// Pools d'objets (docs/04 § 9) : instances déclarées une fois pour toutes, attribuées au déploiement par
// FB_ObjectFactory. La bibliothèque fournit FB_DefaultPools ; un projet peut donner les siens.
INTERFACE I_ObjectPools

// Nombre d'éléments du pool d'un type, 0 = type absent
METHOD PoolSize : UINT
VAR_INPUT
    nType : UINT;
END_VAR
END_METHOD

// N° du pool d'un type : deux types qui partagent un pool (axe linéaire et rotatif, modules) ont le même n°
METHOD PoolId : UINT
VAR_INPUT
    nType : UINT;
END_VAR
END_METHOD

// Élément nIndex (1..PoolSize) du pool d'un type
METHOD Element : I_Object
VAR_INPUT
    nType : UINT;
    nIndex : UINT;
END_VAR
END_METHOD

END_INTERFACE

(* stored: Version 1.1.0.1, ProductVersion 3.1.4024.12
   Itf I_ObjectPools: Id {e3a6014a-d26d-5d26-9218-d619834af91f}
   Method PoolSize: Id {888f9d33-7137-502f-8d7b-b3bbf14089a3}
   Method PoolId: Id {8bae74f9-df38-5424-b4c6-964c7c87ba5a}
   Method Element: Id {3b21351e-821d-5cc2-99b8-5f44f9ff9eb7} *)
